INTERFACE I_Message EXTENDS I_CatalogEvent

METHOD Send : HRESULT
END_METHOD

END_INTERFACE

(* stored: Version 1.1.0.1, ProductVersion 3.1.4026.26
   Itf I_Message: Id {93f0d335-f913-4849-8ca7-510ba6ea7fe4}
   Method Send: Id {7abe0bd7-d420-47c1-99b2-a35bd7343479} *)
